// TIA Portal V20 export
// export: Created 2026-10-20T18:54:53.8019093Z, ExportSetting None, DisplayName Totally Integrated Automation Portal, DisplayVersion V20 Update 6, DisplayName TIA Portal Openness, DisplayVersion V20 Update 6, DisplayName TIA Portal Version Control Interface, DisplayVersion V20 Update 6, DisplayName SINAMICS Startdrive Advanced, DisplayVersion V20 SP1, DisplayName SINAMICS Startdrive G130, G150, S120, S150, SINAMICS MV, G220, S200, S210, DisplayVersion V20 SP1, DisplayName SINAMICS Startdrive G110M, G120, G120C, G120D, G120P, G115D, DisplayVersion V20 SP1, DisplayName STEP 7 Professional, DisplayVersion V20 Update 6, DisplayName STEP 7 Safety, DisplayVersion V20 Update 2, DisplayName WinCC Basic/Comfort/Advanced, DisplayVersion V20 Update 6, DisplayName WinCC Unified, DisplayVersion V20 Update 6
VAR_GLOBAL   // PLC tag table "IO_VFDs_2"
   VTD2_ControlWord AT %QW216 : Word;
   VTD2_MainSetpoint AT %QW218 : Word;
   VTD2_ActualSpeed AT %IW488 : Word;
   VTD2_ActualCurrent AT %IW490 : Word;
   C2101_ControlWord AT %QW224 : Word;
   C2101_MainSetpoint AT %QW226 : Word;
   C2101_StatusWord AT %IW2222 : Word;
   C2101_ActualSpeed AT %IW2224 : Word;
   C2101_ActualCurrent AT %IW2226 : Word;
   C2102_ControlWord AT %QW228 : Word;
   C2102_MainSetpoint AT %QW230 : Word;
   C2102_StatusWord AT %IW2234 : Word;
   C2102_ActualSpeed AT %IW2236 : Word;
   C2102_ActualCurrent AT %IW2238 : Word;
   C2103_ControlWord AT %QW232 : Word;
   C2103_MainSetpoint AT %QW234 : Word;
   C2103_StatusWord AT %IW2246 : Word;
   C2103_ActualSpeed AT %IW2248 : Word;
   C2103_ActualCurrent AT %IW2250 : Word;
   C2104_ControlWord AT %QW308 : Word;
   C2104_MainSetpoint AT %QW310 : Word;
   C2104_StatusWord AT %IW2258 : Word;
   C2104_ActualSpeed AT %IW2260 : Word;
   C2104_ActualCurrent AT %IW2262 : Word;
   C2105_ControlWord AT %QW325 : Word;
   C2105_MainSetpoint AT %QW327 : Word;
   C2105_StatusWord AT %IW2294 : Word;
   C2105_ActualSpeed AT %IW2296 : Word;
   C2105_ActualCurrent AT %IW2298 : Word;
   C2106_ControlWord AT %QW312 : Word;
   C2106_MainSetpoint AT %QW314 : Word;
   C2106_StatusWord AT %IW2270 : Word;
   C2106_ActualSpeed AT %IW2272 : Word;
   C2106_ActualCurrent AT %IW2274 : Word;
   C2107_ControlWord AT %QW316 : Word;
   C2107_MainSetpoint AT %QW318 : Word;
   C2107_StatusWord AT %IW2282 : Word;
   C2107_ActualSpeed AT %IW2284 : Word;
   C2107_ActualCurrent AT %IW2286 : Word;
   CVTD2_ControlWord AT %QW220 : Word;
   CVTD2_MainSetpoint AT %QW222 : Word;
   CVTD2_StatusWord AT %IW2210 : Word;
   CVTD2_ActualSpeed AT %IW2212 : Word;
   CVTD2_ActualCurrent AT %IW2214 : Word;
   C2108_ControlWord AT %QW334 : Word;
   C2108_MainSetpoint AT %QW336 : Word;
   C2108_StatusWord AT %IW2306 : Word;
   C2108_ActualSpeed AT %IW2308 : Word;
   C2108_ActualCurrent AT %IW2310 : Word;
   C2201_ActualCurrent AT %IW2322 : Word;
   C2201_ActualSpeed AT %IW2320 : Word;
   C2201_ControlWord AT %QW338 : Word;
   C2201_MainSetpoint AT %QW340 : Word;
   C2201_StatusWord AT %IW2318 : Word;
   C2202_ActualCurrent AT %IW2334 : Word;
   C2202_ActualSpeed AT %IW2332 : Word;
   C2202_ControlWord AT %QW342 : Word;
   C2202_MainSetpoint AT %QW344 : Word;
   C2202_StatusWord AT %IW2330 : Word;
   C2203_ActualCurrent AT %IW2346 : Word;
   C2203_ActualSpeed AT %IW2344 : Word;
   C2203_ControlWord AT %QW346 : Word;
   C2203_MainSetpoint AT %QW348 : Word;
   C2203_StatusWord AT %IW2342 : Word;
   C2204_ActualCurrent AT %IW2358 : Word;
   C2204_ActualSpeed AT %IW2356 : Word;
   C2204_ControlWord AT %QW351 : Word;
   C2204_MainSetpoint AT %QW353 : Word;
   C2204_StatusWord AT %IW2354 : Word;
   C2205_ActualCurrent AT %IW2370 : Word;
   C2205_ActualSpeed AT %IW2368 : Word;
   C2205_ControlWord AT %QW355 : Word;
   C2205_MainSetpoint AT %QW357 : Word;
   C2205_StatusWord AT %IW2366 : Word;
   C2206_ActualCurrent AT %IW2382 : Word;
   C2206_ActualSpeed AT %IW2380 : Word;
   C2206_ControlWord AT %QW359 : Word;
   C2206_MainSetpoint AT %QW361 : Word;
   C2206_StatusWord AT %IW2378 : Word;
   C2207_ActualCurrent AT %IW2394 : Word;
   C2207_ActualSpeed AT %IW2392 : Word;
   C2207_ControlWord AT %QW363 : Word;
   C2207_MainSetpoint AT %QW365 : Word;
   C2207_StatusWord AT %IW2390 : Word;
   C2208_ActualCurrent AT %IW2406 : Word;
   C2208_ActualSpeed AT %IW2404 : Word;
   C2208_ControlWord AT %QW472 : Word;
   C2208_MainSetpoint AT %QW474 : Word;
   C2208_StatusWord AT %IW2402 : Word;
   VTD2_StatusWord AT %IW486 : Word;
   VTD2_ActualTorque AT %IW492 : Word;
   C2207_ActualTorque AT %IW2396 : Word;
   C2208_ActualTorque AT %IW2408 : Word;
   C2203_ActualTorque AT %IW2348 : Word;
   C2104_ActualTorque AT %IW2264 : Word;
   C2106_ActualTorque AT %IW2276 : Word;
   C2201_ActualTorque AT %IW2324 : Word;
   C2205_ActualTorque AT %IW2372 : Word;
   C2204_ActualTorque AT %IW2360 : Word;
   C2206_ActualTorque AT %IW2384 : Word;
   C2202_ActualTorque AT %IW2336 : Word;
   CVTD2_ActualTorque AT %IW2216 : Word;
   C2103_ActualTorque AT %IW2252 : Word;
   C2107_ActualTorque AT %IW2288 : Word;
   C2105_ActualTorque AT %IW2300 : Word;
   C2102_ActualTorque AT %IW2240 : Word;
   C2101_ActualTorque AT %IW2228 : Word;
   C2108_ActualTorque AT %IW2312 : Word;
   VTD2_AccFactor AT %QW1517 : Word;
END_VAR
